(* IEC 61131-3 sources: Gen-AI/docs/member2_validation/codesys_release_v1.1/C02_type, 1 file *)

(* ---- source.st ---- *)
FUNCTION_BLOCK FB_AgentProbeType
VAR_OUTPUT
 y : BOOL;
END_VAR
y := 'not-a-bool';
END_FUNCTION_BLOCK
